(*
SPDX-FileCopyrightText: © 2026 Oleksandr Tiutyk <trofimich@gmail.com>
SPDX-License-Identifier: MIT
License: https://opensource.org/license/mit
*)

(*!
<summary>Runs one automation component scenario in an isolated fixture.</summary>
<description>
Owns a freshly allocated fixture for the active run. AfterTest releases it after success or a reported
exception. A concrete pointer preserves FB_exit for the fixture and its nested resource owners.
Use one task. Do not copy the test case while it owns a fixture.
</description>
*)

{attribute 'no_assign'}
{attribute 'no_explicit_call' := 'do not call this function block directly'}
FUNCTION_BLOCK AutomationComponentTestCase EXTENDS TOF_Testing.SingleCycleTest
VAR_STAT
	{attribute 'hide'}
	_ClassName : STRING := __POUNAME();
END_VAR
VAR
	_Scenario : AUTOMATION_COMPONENT_TEST_SCENARIO;
	_Fixture : POINTER TO AutomationComponentTestFixture;
END_VAR

(*!
<summary>Selects the scenario without allocating its fixture.</summary>
<param name="name">Name reported for this case.</param>
<param name="parent">Group that owns this case.</param>
<param name="scenario">Scenario selected for the case.</param>
*)
METHOD FB_init : BOOL
VAR_INPUT
	bInitRetains: BOOL; // TRUE: the retain variables are initialized (reset warm / reset cold)
	bInCopyCode: BOOL; // TRUE: the instance will be copied to the copy code afterward (online change)
	name : WSTRING;
	parent : TOF_Testing.ITestElement;
	scenario : AUTOMATION_COMPONENT_TEST_SCENARIO;
END_VAR
IF NOT bInCopyCode THEN
	_Scenario := scenario;
END_IF

FB_init := TRUE;
END_METHOD

(*!
<summary>Allocates a fresh fixture and runs the selected scenario.</summary>
<description>Terminal allocation failure is raised at the task boundary after case handling.</description>
*)
METHOD PROTECTED ExecuteTest
VAR
	assertions : REFERENCE TO TOF_Testing.Assertions;
END_VAR
_Fixture := __NEW(AutomationComponentTestFixture);

IF _Fixture = 0 THEN
	TOF_Core.DynamicMemoryManager.RaiseAllocationFailure();

	RETURN;
END_IF

assertions REF= Assert;
_Fixture^.ExecuteScenario(scenario := _Scenario, assertions := assertions);
END_METHOD

(*!
<summary>Releases the fixture before the case outcome is published.</summary>
<description>The framework records an exception from teardown. Clear the stored alias before releasing.</description>
*)
METHOD PROTECTED AfterTest
VAR
	fixture : POINTER TO AutomationComponentTestFixture;
END_VAR
fixture := _Fixture;
_Fixture := 0;

IF fixture <> 0 THEN
	__DELETE(fixture);
END_IF
END_METHOD

(*!
<summary>Releases an active fixture if the case is unloaded before its teardown.</summary>
<description>The fixture and its nested FB_exit paths complete without exceptions.</description>
<param name="bInCopyCode">TwinCAT copy-code exit marker. The previous instance leaves copied storage alive.</param>
*)
METHOD FB_exit : BOOL
VAR_INPUT
	bInCopyCode : BOOL;
END_VAR
IF NOT bInCopyCode AND_THEN _Fixture <> 0 THEN
	__DELETE(_Fixture);
END_IF

FB_exit := TRUE;
END_METHOD

(*!
<summary>Borrows the concrete class name. Callers must not modify it.</summary>
*)
{attribute 'monitoring' := 'call'}
PROPERTY ClassName : REFERENCE TO STRING
GET
ClassName REF= _ClassName;
END_GET
END_PROPERTY

(*!
<summary>Borrows the project namespace name. Callers must not modify it.</summary>
*)
{attribute 'monitoring' := 'call'}
PROPERTY NamespaceName : REFERENCE TO STRING
GET
NamespaceName REF= CurrentNamespace.Name;
END_GET
END_PROPERTY

(*!
<summary>Reports the complete instance size in bytes.</summary>
*)
{attribute 'monitoring' := 'call'}
PROPERTY SelfSize : ULINT
GET
SelfSize := XSIZEOF(THIS^);
END_GET
END_PROPERTY

END_FUNCTION_BLOCK

(* stored: Version 1.1.0.1
   POU AutomationComponentTestCase: Id {539ed20f-c987-435d-9bc2-50e3d6d452cb}, SpecialFunc None
   Method FB_init: Id {e21bea5d-f495-47c0-8255-c4844a55b2e9}
   Method ExecuteTest: Id {99754db6-5e4b-4d56-86e1-06a9b2f21d9e}
   Method AfterTest: Id {ac04e650-5217-47d3-bb37-48d9ced549f7}
   Method FB_exit: Id {b6ee1d00-7204-4014-884c-6174651a21d2}
   Property ClassName: Id {e5db47dd-42dc-4a03-8151-11003399d67e}
   Get Get: Id {2c22e41b-c2e4-4189-8de1-bf27f15015b7}
   Property NamespaceName: Id {181278a1-326d-4093-8bc7-7cb2a6f794c1}
   Get Get: Id {40c813c7-abcd-4b7a-885d-6ea816dbc553}
   Property SelfSize: Id {9b7ac916-61a6-442a-a149-63e5d5630f02}
   Get Get: Id {345469e4-faaf-4525-a916-08abb7961f8e} *)
